(* IEC 61131-3 sources: llm-plc-st-eval/data/definitivo/qwen2.5-coder_14b/I2/zero_shot, 3 files *)

(* ---- ejec_1.st ---- *)
```pascal
FUNCTION_BLOCK FB_Llenado
VAR_INPUT
    nivelAlto, nivelBajo, btnInicio, btnParo : BOOL;
END_VAR

VAR_OUTPUT
    vLlenado, motorMezcla, vDescarga : BOOL;
END_VAR

VAR
    estado : INT := 0; // 0: reposo, 1: llenado, 2: mezcla, 3: descarga
    timerMezcla : TON;
END_VAR

// Estado de reposo
IF btnParo THEN
    estado := 0;
    vLlenado := FALSE;
    motorMezcla := FALSE;
    vDescarga := FALSE;
    timerMezcla(IN := FALSE);
ELSIF btnInicio AND estado = 0 THEN
    estado := 1;
    vLlenado := TRUE;
END_IF

// Estado de llenado
IF estado = 1 THEN
    IF nivelAlto THEN
        estado := 2;
        vLlenado := FALSE;
        motorMezcla := TRUE;
        timerMezcla(IN := TRUE, PT := T#60S);
    END_IF
END_IF

// Estado de mezcla
IF estado = 2 THEN
    IF timerMezcla.Q THEN
        estado := 3;
        motorMezcla := FALSE;
        vDescarga := TRUE;
    END_IF
END_IF

// Estado de descarga
IF estado = 3 THEN
    IF nivelBajo THEN
        estado := 0;
        vDescarga := FALSE;
    END_IF
END_IF
```

Este código implementa un proceso de llenado por etapas utilizando un FUNCTION_BLOCK en Structured Text (ST) conforme al estándar IEC 61131-3. Las variables de entrada y salida están declaradas al principio, y se utiliza un temporizador (`timerMezcla`) para controlar la duración de la mezcla. El proceso se puede detener en cualquier momento con el botón `btnParo`, llevando todas las salidas a un estado seguro.

(* ---- ejec_2.st ---- *)
```pascal
FUNCTION_BLOCK FB_Llenado
VAR_INPUT
    nivelAlto : BOOL;  // Nivel alto detectado
    nivelBajo : BOOL;  // Nivel bajo detectado
    btnInicio : BOOL;  // Botón de inicio
    btnParo   : BOOL;  // Botón de paro
END_VAR

VAR_OUTPUT
    vLlenado  : BOOL;  // Válvula de llenado
    motorMezcla : BOOL;  // Motor de mezcla
    vDescarga : BOOL;  // Válvula de descarga
END_VAR

VAR
    estado : INT := 0;  // Estado actual del proceso
    timerMezcla : TON;  // Timer para el motor de mezcla
END_VAR

// Inicialización del timer
timerMezcla(IN := FALSE, PT := T#60S);

// Máquina de estados
CASE estado OF
    0:  // Reposo
        IF btnInicio THEN
            estado := 1;  // Iniciar el proceso de llenado
        END_IF;
    1:  // Llenado
        vLlenado := TRUE;
        IF nivelAlto THEN
            estado := 2;  // Pasar al siguiente estado después de alcanzar el nivel alto
        END_IF;
    2:  // Mezcla
        vLlenado := FALSE;
        motorMezcla := TRUE;
        timerMezcla(IN := TRUE);
        IF timerMezcla.Q THEN
            estado := 3;  // Pasar al siguiente estado después de 60 segundos
        END_IF;
    3:  // Descarga
        motorMezcla := FALSE;
        vDescarga := TRUE;
        IF nivelBajo THEN
            estado := 0;  // Regresar al reposo después de alcanzar el nivel bajo
        END_IF;
END_CASE;

// Manejo del botón de paro
IF btnParo THEN
    estado := 0;  // Regresar al reposo
    vLlenado := FALSE;
    motorMezcla := FALSE;
    vDescarga := FALSE;
    timerMezcla(IN := FALSE);  // Detener el timer
END_IF;
```

Este código implementa una máquina de estados para controlar un proceso de llenado por etapas utilizando un FUNCTION_BLOCK en Structured Text (ST) conforme al estándar IEC 61131-3. El proceso pasa por las etapas de llenado, mezcla y descarga, y puede ser detenido en cualquier momento mediante el botón de paro, llevando todas las salidas a un estado seguro.

(* ---- ejec_3.st ---- *)
```iec
FUNCTION_BLOCK FB_Llenado
VAR_INPUT
    nivelAlto : BOOL; // Nivel alto detectado
    nivelBajo : BOOL; // Nivel bajo detectado
    btnInicio : BOOL; // Botón de inicio
    btnParo : BOOL; // Botón de paro
END_VAR

VAR_OUTPUT
    vLlenado : BOOL; // Válvula de llenado
    motorMezcla : BOOL; // Motor de mezcla
    vDescarga : BOOL; // Válvula de descarga
END_VAR

VAR
    estado : INT := 0; // Estado actual del proceso
    timerMezcla : TON; // Timer para el motor de mezcla
    timerMezclaPT : TIME := T#60S; // Periodo de tiempo para el motor de mezcla
END_VAR

// Inicialización del timer
timerMezcla(IN := FALSE, PT := timerMezclaPT);

// Máquina de estados
CASE estado OF
    0: // Reposo
        vLlenado := FALSE;
        motorMezcla := FALSE;
        vDescarga := FALSE;
        IF btnInicio THEN
            estado := 1; // Iniciar el llenado
        END_IF;
        IF btnParo THEN
            estado := 0; // Mantener en reposo si se presiona btnParo
        END_IF;

    1: // Llenado
        vLlenado := TRUE;
        motorMezcla := FALSE;
        vDescarga := FALSE;
        IF nivelAlto THEN
            estado := 2; // Pasar al siguiente estado después de alcanzar nivel alto
        END_IF;
        IF btnParo THEN
            estado := 0; // Parar el proceso si se presiona btnParo
        END_IF;

    2: // Mezcla
        vLlenado := FALSE;
        motorMezcla := TRUE;
        vDescarga := FALSE;
        timerMezcla(IN := TRUE);
        IF timerMezcla.Q THEN
            estado := 3; // Pasar al siguiente estado después de 60 segundos
        END_IF;
        IF btnParo THEN
            estado := 0; // Parar el proceso si se presiona btnParo
        END_IF;

    3: // Descarga
        vLlenado := FALSE;
        motorMezcla := FALSE;
        vDescarga := TRUE;
        IF nivelBajo THEN
            estado := 0; // Regresar a reposo después de alcanzar nivel bajo
        END_IF;
        IF btnParo THEN
            estado := 0; // Parar el proceso si se presiona btnParo
        END_IF;

    ELSE
        estado := 0; // Mantener en reposo si el estado no está definido
END_CASE;
```

Este código implementa una máquina de estados para controlar un proceso de llenado por etapas utilizando un FUNCTION_BLOCK en Structured Text (ST) conforme al estándar IEC 61131-3. Las variables de entrada y salida están declaradas y se utilizan para controlar las etapas del proceso. El botón de paro detiene el proceso y regresa a un estado seguro.
